Fanuc KAREL source: kt00452.KL

-- PROVISIONAL review KL for V1013-1; original PC SHA256 0e7fb6a9623c9b5078723d9ea1b7dba9877ed88e47659f0777bd15994d1f3f25
-- Incomplete behavior may be omitted. Consult companion uncertainty JSON. Do not deploy.
PROGRAM KT00452
%NOLOCKGROUP
VAR
  R2 : REAL
  OUT : BOOLEAN
-- UNRESOLVED_DECL H1 type=002017
BEGIN
  -- UNRESOLVED_PC offsets 5-19; opcodes 2E,22,9D,33,B4
  -- UNRESOLVED_PC offsets 24-35; opcodes 2E,23
  -- UNRESOLVED_PC offsets 40-65; opcodes 22,9D,33,B3,21,29,64,29,72,23
  -- UNRESOLVED_PC offsets 70-74; opcodes 7F
END KT00452
